ABB RobotStudio station: gofa_chess.rspag

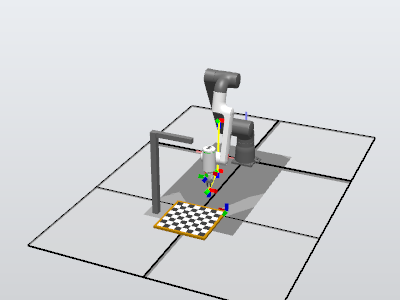
--- station ---
Station gofa_real_accurate (saved by RobotStudio 26.2.11700.0)
Controller Controller2
  mechanical unit ROB_1: CRB15000_10_152__01, 6 joints, base frame (0, 0, 0) mm
Layout (positions relative to the parent item):
  - CRB15000_10_152__01 [mechanism, from %ABB.RobotStudio.Models.CRB15000%\CRB15000_10_152__01.rslib] at (0, 0, 0) mm; joint values [1.5933, 0.5665, 0.7265, 0, 0.2778, 1.5933] (rad or m)
  - surface_1 [part], size 410 x 1236 x 0 mm
  - surface_4 [part], size 374 x 1236 x 0 mm
  - surface_3 [part], size 374 x 258 x 0 mm
  - surface_2 [part], size 410 x 258 x 0 mm
  - chess_board [part] at (0, 1209.66, 30) mm, size 440 x 440 x 20 mm
  - Smart_Gripper_Servo_Fingers [mechanism, from %ABB.RobotStudio.Models.SmartGripper%\ABB_Smart_Gripper_Servo_Fingers.rslib] at (-20, 889.66, 313.14) mm, rotated rx -180 ry 0 rz 180 deg; joint values [0.0102] (rad or m)
  - PoseMover [smart component, from Components\PoseMover.rslib]
      properties: Mechanism=Smart_Gripper_Servo_Fingers; Pose=3; Duration=0
  - PoseMover_2 [smart component, from Components\PoseMover.rslib]
      properties: Mechanism=Smart_Gripper_Servo_Fingers; Pose=2; Duration=0
  - LogicGate [smart component, from Components\LogicGate.rslib]
      properties: Operator=NOT; Delay=0
  - Part_1 [part] at (354.61, 1137.15, 0) mm, size 50 x 50 x 730 mm
  - Part_2 [part], size 300 x 40 x 40 mm
Attachment: Smart_Gripper_Servo_Fingers is attached to CRB15000_10_152__01 / Link6
Station logic (signal -> signal, property => property):
  LogicGate.Output -> PoseMover_2.Execute
  Controller2.DO_Gripper -> LogicGate.InputA
  Controller2.DO_Gripper -> PoseMover.Execute

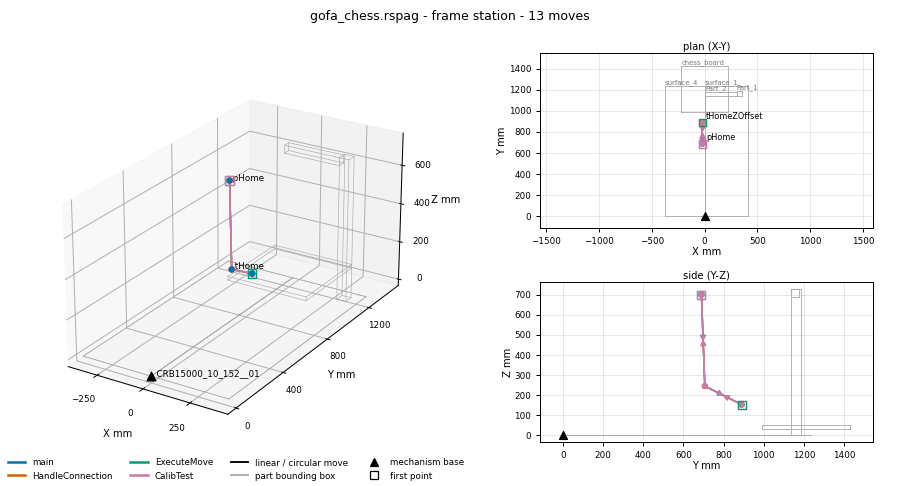
[picture p0: tool path of gofa_chess.rspag in frame station, 13 of 16 moves have a stored position in this frame; points joined in program order, loops and branches not executed]
--- Controller Data/Controller2/RAPID/TASK2/PROGMOD/CalibData.modx ---
MODULE CalibData
    PERS tooldata Camera:=[TRUE,[[-7.3,28.3,35.1],[0.5,-0.5,0.5,0.5]],[0.229,[7.9,12.4,48.7],[1,0,0,0],0.00021,0.00023,0.00008]];
    !PERS tooldata Servo:=[TRUE,[[0,0,114.2],[1,0,0,0]],[0.215,[8.7,12.3,49.2],[1,0,0,0],0.00021,0.00024,0.00009]];
    !TASK PERS wobjdata chess_workobj:=[FALSE,TRUE,"",[[0,0,0],[1,0,0,0]],[[-220,580,420],[1,0,0,0]]];
ENDMODULE

--- Controller Data/Controller2/RAPID/TASK2/PROGMOD/ChessMotion.modx ---
MODULE ChessMotion
    ! Socket Variables
    VAR socketdev server_socket;
    VAR socketdev client_socket;
    VAR string received_cmd;

    ! Array to hold [Action, X, Y] sent from Python
    ! Action: 1 = PICK, 2 = PLACE
    VAR num cmd_data{3};
    VAR bool is_parsed;

    ! --- TOOL AND WORKOBJECT DEFINITIONS ---
    PERS tooldata Servo:=[TRUE,[[0,0,160],[1,0,0,0]],[0.215,[8.7,12.3,49.2],[1,0,0,0],0.00021,0.00024,0.00009]];
    TASK PERS wobjdata chess_workobj:=[FALSE,TRUE,"",[[0,0,0],[1,0,0,0]],[[-220,989.663,50],[1,0,0,0]]];

    ! --- HOME POSITION ---
    ! Defines a safe parking spot 250mm above the center-ish of the board
    CONST robtarget pHome := [[200,-300,650],[0,0,1,0],[0,0,0,0],[9E+09,9E+09,9E+09,9E+09,9E+09,9E+09]];
    CONST robtarget tHome := [[200,-283.240199578,195.507235305],[0,0,1,0],[0,0,0,0],[9E+09,9E+09,9E+09,9E+09,9E+09,9E+09]];
    CONST robtarget tHomeZOffset := [[199.999965031,-100.000072343,103.135393127],[-0,0,1,-0.000000014],[1,-1,1,0],[9E+09,9E+09,9E+09,9E+09,9E+09,9E+09]];

    PROC main()
        ! 1. SAFE STARTUP SEQUENCE
!        SetDO DO_Gripper, 0;  ! Ensure gripper is physically OPEN at startup
        PulseDO\PLength:=0.2,DO16_GripperOpen;
        WaitTime 0.5;

        ! Move safely to the Home position before accepting any commands
        ! Using MoveJ (Joint move) to avoid singularity/linear path errors from unknown start poses
        MoveJ pHome, v200, z10, Servo \WObj:=chess_workobj;
        MoveL tHome, v200, z10, Servo \WObj:=chess_workobj;
        MoveL tHomeZOffset, v200, fine, Servo \WObj:=chess_workobj;

        ! 2. START SERVER
        SocketCreate server_socket;
        SocketBind server_socket, "127.0.0.1", 5000;
        SocketListen server_socket;

        WHILE TRUE DO
            TPWrite "Waiting for Python on port 5000...";
            SocketAccept server_socket, client_socket;
            HandleConnection;
            SocketClose client_socket;
        ENDWHILE
    ENDPROC

    PROC HandleConnection()
        WHILE TRUE DO
            ! Added \Time:=WAIT_MAX so the robot waits forever while you think
            SocketReceive client_socket \Str:=received_cmd \Time:=WAIT_MAX;

            ! Instantly convert string "[1, 200, 150]" into the cmd_data array
            is_parsed := StrToVal(received_cmd, cmd_data);

            IF is_parsed THEN
                ! Call our dynamic macro using the parsed X (cmd_data{2}) and Y (cmd_data{3})
                ExecuteMove cmd_data{1}, cmd_data{2}, cmd_data{3};
                SocketSend client_socket \Str:="DONE";
            ELSE
                TPWrite "Error: Bad format -> " + received_cmd;
                SocketSend client_socket \Str:="ERROR";
            ENDIF
        ENDWHILE
    ERROR
        ! If a timeout error still somehow occurs, just ignore it and wait again
        IF ERRNO = ERR_SOCK_TIMEOUT THEN
            RETRY;
        ENDIF

        TPWrite "Python disconnected.";

        ! Park safely back at home when the game/script ends
        ! Using MoveL to safely back out of the camera's L-bracket structure linearly
        MoveL tHomeZOffset, v200, z10, Servo \WObj:=chess_workobj;
        MoveL tHome, v200, z10, Servo \WObj:=chess_workobj;
        MoveL pHome, v200, z10, Servo \WObj:=chess_workobj;

        RETURN;
    ENDPROC

    ! --- THE DYNAMIC PICK AND PLACE MACRO ---
    PROC ExecuteMove(num action, num target_x, num target_y)
        ! 1. ALL variables must be declared at the very top
        VAR robtarget base_target;
        VAR num hover_height := 100; ! Hover 100mm above the piece

        ! --- Z OFFSET CONTROL ---
        ! Change this value to adjust pickup height.
        ! Positive = Higher up, Negative = Deeper down.
        VAR num z_offset := 25;

        ! 2. NOW executable statements can begin
        base_target := [[target_x, target_y, z_offset], [0, 0, 1, 0], [0, 0, 0, 0], [9E9, 9E9, 9E9, 9E9, 9E9, 9E9]];

        ! 3. Approach position (Hover)
        MoveL Offs(base_target, 0, 0, hover_height), v200, z10, Servo \WObj:=chess_workobj;

        ! 4. Move down to the piece
        MoveL base_target, v50, fine, Servo \WObj:=chess_workobj;

        ! 5. Actuate Gripper
        IF action = 1 THEN
!            SetDO DO_Gripper, 1; ! Close gripper (PICK)
            PulseDO\PLength:=0.2,DO16_GripperClose;
            WaitTime 0.5;
        ELSEIF action = 2 THEN
!            SetDO DO_Gripper, 0; ! Open gripper (PLACE)
            PulseDO\PLength:=0.2,DO16_GripperOpen;

            WaitTime 0.5;
        ENDIF

        ! 6. Retract safely back up to hover height
        MoveL Offs(base_target, 0, 0, hover_height), v200, z10, Servo \WObj:=chess_workobj;

        ! 7. Return to the intermediate home position ONLY after a PLACE action
        IF action = 2 THEN
            MoveL tHomeZOffset, v200, z10, Servo \WObj:=chess_workobj;
        ENDIF
    ENDPROC

    PROC CalibTest()
        TPWrite "--- Starting Calibration Dry Run ---";

        ! 1. SAFE STARTUP APPROACH
!        SetDO DO_Gripper, 0; ! Ensure gripper is open
        PulseDO\PLength:=0.2,DO16_GripperOpen;
        WaitTime 0.5;
        MoveJ pHome, v200, z10, Servo \WObj:=chess_workobj;
        MoveL tHome, v200, z10, Servo \WObj:=chess_workobj;
        MoveL tHomeZOffset, v200, fine, Servo \WObj:=chess_workobj;

        ! 2. TEST POINTS (Action 0 = No gripper actuation)
        ! Test Near Corner (approx A1/H1)
        TPWrite "Testing Corner 1 (21, 21)...";
        ExecuteMove 0, 21, 21;

        ! Test Far Corner (approx H8/A8)
        TPWrite "Testing Corner 2 (315, 315)...";
        ExecuteMove 0, 315, 315;

        ! Test Center of Board
        TPWrite "Testing Center (168, 168)...";
        ExecuteMove 0, 168, 168;

        TPWrite "Calibration Complete. Retracting safely...";

        ! 3. SAFE LINEAR RETRACTION (Camera Avoidance)
        MoveL tHomeZOffset, v200, z10, Servo \WObj:=chess_workobj;
        MoveL tHome, v200, z10, Servo \WObj:=chess_workobj;
        MoveL pHome, v200, fine, Servo \WObj:=chess_workobj;

        TPWrite "--- Routine Finished ---";
    ENDPROC

ENDMODULE

--- Controller Data/Controller2/RAPID/TASK2/PROGMOD/Wizard_LoadData.modx ---
MODULE Wizard_LoadData
ENDMODULE

--- Controller Data/Controller2/RAPID/TASK2/SYSMOD/Wizard_Params.sysx ---
MODULE Wizard_Params (SYSMODULE)
    !***************************************************************************
    !*                              Common parameters                          *
    !***************************************************************************
    ! Predefined common targets for user to use
    CONST jointtarget wi_jPosCalib:=[[0,0,0,0,30,0],[9E+9,9E+9,9E+9,9E+9,9E+9,9E+9]];

	PERS robtarget wi_homePosition:=[[597.47,0.00,837.78],[0.5,0,0.866025,0],[0,0,0,0],[9E+9,9E+9,9E+9,9E+9,9E+9,9E+9]];

    VAR errnum wi_errnum;

    PERS bool wi_bFirstLaunched:=TRUE;

    PERS string wi_asiMoveType:="move_to_location";

    ! The parameter is the option sequence of Speed dropdown
    PERS string wi_speed:="VQUICK:v1000,QUICK:v500,MODERATE:v200,SLOW:v50,VSLOW:v20";

    ! This proc is the rapid placeholder for empty procedure filed in Wizard; Do not remove it
    PROC wi_ProcPlaceHolder_Hidden()
    ENDPROC

ENDMODULE

--- Controller Data/Controller2/HOME/Wizard/Wizard.mod ---
MODULE Wizard
	PROC main()
		<SMT>
	ENDPROC
ENDMODULE

--- Controller Data/Controller2/SYSPAR/EIO.cfg ---
EIO:CFG_1.0:8:0::
#
VIRTUAL_NETWORK:

      -Name "Virtual" -Label "Virtual Device Network"
#
EIO_SIGNAL:

      -Name "IIO_di1" -SignalType "DI" -Device "IntegratedIOInternalDevice"\
      -DeviceMap "0"

      -Name "IIO_di2" -SignalType "DI" -Device "IntegratedIOInternalDevice"\
      -DeviceMap "1"

      -Name "IIO_di3" -SignalType "DI" -Device "IntegratedIOInternalDevice"\
      -DeviceMap "2"

      -Name "IIO_di4" -SignalType "DI" -Device "IntegratedIOInternalDevice"\
      -DeviceMap "3"

      -Name "IIO_di5" -SignalType "DI" -Device "IntegratedIOInternalDevice"\
      -DeviceMap "4"

      -Name "IIO_di6" -SignalType "DI" -Device "IntegratedIOInternalDevice"\
      -DeviceMap "5"

      -Name "IIO_di7" -SignalType "DI" -Device "IntegratedIOInternalDevice"\
      -DeviceMap "6"

      -Name "IIO_di8" -SignalType "DI" -Device "IntegratedIOInternalDevice"\
      -DeviceMap "7"

      -Name "IIO_di9" -SignalType "DI" -Device "IntegratedIOInternalDevice"\
      -DeviceMap "8"

      -Name "IIO_di10" -SignalType "DI" -Device "IntegratedIOInternalDevice"\
      -DeviceMap "9"

      -Name "IIO_di11" -SignalType "DI" -Device "IntegratedIOInternalDevice"\
      -DeviceMap "10"

      -Name "IIO_di12" -SignalType "DI" -Device "IntegratedIOInternalDevice"\
      -DeviceMap "11"

      -Name "IIO_di13" -SignalType "DI" -Device "IntegratedIOInternalDevice"\
      -DeviceMap "12"

      -Name "IIO_di14" -SignalType "DI" -Device "IntegratedIOInternalDevice"\
      -DeviceMap "13"

      -Name "IIO_di15" -SignalType "DI" -Device "IntegratedIOInternalDevice"\
      -DeviceMap "14"

      -Name "IIO_di16" -SignalType "DI" -Device "IntegratedIOInternalDevice"\
      -DeviceMap "15"

      -Name "IIO_do1" -SignalType "DO" -Device "IntegratedIOInternalDevice"\
      -DeviceMap "0"

      -Name "IIO_do2" -SignalType "DO" -Device "IntegratedIOInternalDevice"\
      -DeviceMap "1"

      -Name "IIO_do3" -SignalType "DO" -Device "IntegratedIOInternalDevice"\
      -DeviceMap "2"

      -Name "IIO_do4" -SignalType "DO" -Device "IntegratedIOInternalDevice"\
      -DeviceMap "3"

      -Name "IIO_do5" -SignalType "DO" -Device "IntegratedIOInternalDevice"\
      -DeviceMap "4"

      -Name "IIO_do6" -SignalType "DO" -Device "IntegratedIOInternalDevice"\
      -DeviceMap "5"

      -Name "IIO_do7" -SignalType "DO" -Device "IntegratedIOInternalDevice"\
      -DeviceMap "6"

      -Name "IIO_do8" -SignalType "DO" -Device "IntegratedIOInternalDevice"\
      -DeviceMap "7"

      -Name "IIO_gi" -SignalType "GI" -Device "integratedIOInternalDevice"\
      -DeviceMap "0-15"

      -Name "IIO_go" -SignalType "GO" -Device "integratedIOInternalDevice"\
      -DeviceMap "0-7"

      -Name "DO_Gripper" -SignalType "DO"

      -Name "DO16_GripperClose" -SignalType "DO"

      -Name "DO16_GripperOpen" -SignalType "DO"

#CTRL_SIGNATURE:90VkNvpn/wi3TA64bs0ZwY7L60b4tE9T8oBrTjHeOsoqgbYSuXEZJ03ZlCJ1bIjoNp8Pjq4EOeIeO2A8KgUSDg==

--- Controller Data/Controller2/SYSPAR/PROC.cfg ---
PROC:CFG_1.0:8:0::

#CTRL_SIGNATURE:0h+CoyQnbB4hTaJXDmuzS1X0uNi641WJcpigYcKMIlBsq50ulETkbCJ6TRNDagLjHqQr3kbJbwI3pqitwwAMfg==
